Yaskawa INFORM job: ONCHAMF.JBI

/JOB
//NAME ONCHAMF
//POS
///NPOS 0,0,0,0,0,0
//INST
///DATE 2026/10/26 01:19
///COMM Generated using RoboDK
///ATTR SC,RW
///GROUP1 RB1
NOP
CALL JOB:HOME_KU
END
